(* IEC 61131-3 sources: codesys-ai-industrial-robot-control/plc/src/Process/FB_PickSequence, 3 files *)

(* ---- NextStep.st ---- *)
METHOD PRIVATE NextStep
VAR_INPUT
    eNew : E_PickStep;
END_VAR

eStep := eNew;
xRequested := FALSE;
tonRelease(IN := FALSE);

(* ---- Request.st ---- *)
// Requests a robot command once per step; the handshake in the body executes it.
METHOD PRIVATE Request
VAR_INPUT
    eCmd : E_RobotCmd;
    stTgt : SMC_POS_REF;
END_VAR

IF NOT xRequested AND iCmdPhase = 0 THEN
    eReqCmd := eCmd;
    stReqTarget := stTgt;
    iCmdPhase := 1;
    xRequested := TRUE;
END_IF

(* ---- TrackedPose.st ---- *)
// Pose above the tracked part (PCS_1 origin) at height lrZ, tool pointing down.
METHOD PRIVATE TrackedPose : SMC_POS_REF
VAR_INPUT
    lrZ : LREAL;
END_VAR

TrackedPose.c.X := 0;
TrackedPose.c.Y := 0;
TrackedPose.c.Z := lrZ;
TrackedPose.c.A := GVL_CellGeometry.TOOL_DOWN_A;
TrackedPose.c.B := GVL_CellGeometry.TOOL_DOWN_B;
TrackedPose.c.C := GVL_CellGeometry.TOOL_DOWN_C;
